// TIA Portal V21 export
// export: Created 2026-10-12T11:32:17.1501459Z, ExportSetting WithDefaults, DisplayName Totally Integrated Automation Portal, DisplayVersion V21, DisplayName STEP 7 Professional, DisplayVersion V21, DisplayName STEP 7 Safety, DisplayVersion V21, DisplayName Tech WebApplication, DisplayVersion V21, DisplayName WinCC Basic/Comfort/Advanced, DisplayVersion V21, DisplayName WinCC Unified, DisplayVersion V21
VAR_GLOBAL   // PLC tag table "Default tag table"
   System_Byte AT %MB1 : Byte;
   FirstScan AT %M1.0 : Bool;
   DiagStatusUpdate AT %M1.1 : Bool;
   AlwaysTRUE AT %M1.2 : Bool;
   AlwaysFALSE AT %M1.3 : Bool;
   Clock_Byte AT %MB0 : Byte;
   Clock_10Hz AT %M0.0 : Bool;
   Clock_5Hz AT %M0.1 : Bool;
   "Clock_2.5Hz" AT %M0.2 : Bool;
   Clock_2Hz AT %M0.3 : Bool;
   "Clock_1.25Hz" AT %M0.4 : Bool;
   Clock_1Hz AT %M0.5 : Bool;
   "Clock_0.625Hz" AT %M0.6 : Bool;
   "Clock_0.5Hz" AT %M0.7 : Bool;
   "CONTROL ON FLAG" AT %M2.0 : Bool;
   "MANUAL MODE SELECTED" AT %M2.1 : Bool;
   "AUTO MODE SELECTED" AT %M2.2 : Bool;
   "FAULT RESET FLAG" AT %M2.3 : Bool;
   "FAULT BIT" AT %M2.4 : Bool;
   "MANUAL CONVEYOR FWD ON FLAG" AT %M2.5 : Bool;
   "MANUAL CONVEYOR REV ON FLAG" AT %M2.6 : Bool;
END_VAR
